Yaskawa INFORM job: SAVETRAJ.JBI

/JOB
//NAME SAVETRAJ
///FOLDERNAME FOLDER003
//POS
///NPOS 0,0,0,0,0,0
//INST
///DATE 2018/09/29 10:10
///ATTR SC,RW
///GROUP1 RB1
NOP
TIMER T=0.50
SET B030 1
TIMER T=0.50
END
